(* IEC 61131-3 sources: Versio-VersionControlSystem/fixtures/projects/RefrigeratorControl/Device/Plc Logic/Application/Library/Alarm/POUs/FB_Alarm/Protected, 1 file *)

(* ---- _M_Protected.st ---- *)
METHOD PROTECTED _M_Protected : BOOL
VAR_INPUT
END_VAR

// --- BEGIN IMPLEMENTATION ---
